FUNCTION_BLOCK GiveWorkpiece (* Composite Function Block Type *)
  (* Standard: 61499-2 *)
  (* Version 0.0, 7/2/2026, template *)
  PACKAGE Main;
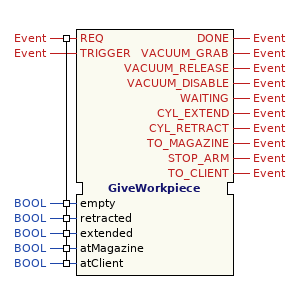
  EVENT_INPUT
    REQ WITH empty, retracted, extended, atMagazine, atClient; (* Normal Execution Request *)
    TRIGGER;
  END_EVENT
  EVENT_OUTPUT
    DONE;
    VACUUM_GRAB;
    VACUUM_RELEASE;
    VACUUM_DISABLE;
    WAITING;
    CYL_EXTEND;
    CYL_RETRACT;
    TO_MAGAZINE;
    STOP_ARM;
    TO_CLIENT;
  END_EVENT
  VAR_INPUT
    empty : BOOL; (* Input event qualifier *)
    retracted : BOOL;
    extended : BOOL;
    atMagazine : BOOL;
    atClient : BOOL;
  END_VAR
  FBS
    FB1 : MagazineSupplyWp;
    ToMagazine : SimpleMove;
    Grab : VacuumSequence;
    ToClient : SimpleMove;
    Release : VacuumSequence;
    FB6 : ArmReset;
    FB7 : E_MERGE;
    FB8 : E_MERGE;
    FB9 : E_MERGE;
    FB10 : E_MERGE;
    FB11 : E_MERGE;
    FB12 : E_MERGE;
  END_FBS
  EVENT_CONNECTIONS
    REQ TO FB1.E7ACA3FA6937DBD5;
    REQ TO ToMagazine.08A6921781769002;
    REQ TO ToClient.08A6921781769002;
    REQ TO FB6.78E8E2AA9DAF29A8;
    TRIGGER TO FB1.CCDC0F1EC03E3A5A;
    FB1.FFF627DF72AA63EC TO CYL_EXTEND;
    FB1.CD1413F90346ACAE TO CYL_RETRACT;
    FB1.F53F7251A3029812 TO ToMagazine.BEEA5224F96B4EAA;
    FB1.C1D84DB1B6EB4247 TO WAITING;
    ToMagazine.19B414802953B8F9 TO Grab.E95F52AEE292CFEA;
    ToMagazine.4A40729E5CEB7782 TO FB11.EI1;
    ToMagazine.FCE01ED48ED44FD9 TO FB12.EI1;
    Grab.8B550AE5A1007C15 TO ToClient.BEEA5224F96B4EAA;
    Grab.5305E856C95E0A15 TO FB7.EI1;
    Grab.2E956B9A6CBDEE5C TO FB8.EI1;
    Grab.993B0E497578A534 TO FB9.EI1;
    ToClient.19B414802953B8F9 TO Release.98EBB230BBACE9D4;
    ToClient.4A40729E5CEB7782 TO FB10.EI1;
    ToClient.FCE01ED48ED44FD9 TO FB12.EI2;
    Release.993B0E497578A534 TO FB9.EI2;
    Release.2E956B9A6CBDEE5C TO FB8.EI2;
    Release.5305E856C95E0A15 TO FB7.EI2;
    Release.8B550AE5A1007C15 TO FB6.44541FA90B36D44F;
    FB6.6B9B16A5CCCF0A5F TO DONE;
    FB6.AF051DE6AC146B46 TO FB10.EI2;
    FB6.88EB222F28F57D09 TO FB11.EI2;
    FB6.4279AF5F2D571F35 TO FB12.EI1;
    FB12.EO TO STOP_ARM;
    FB11.EO TO TO_MAGAZINE;
    FB10.EO TO TO_CLIENT;
    FB9.EO TO VACUUM_DISABLE;
    FB8.EO TO VACUUM_RELEASE;
    FB7.EO TO VACUUM_GRAB;
  END_CONNECTIONS
  DATA_CONNECTIONS
    empty TO FB1.65B96A6108347471;
    retracted TO FB1.F3A16FF43FB1E09C;
    extended TO FB1.F24DAEB350B1D1C4;
    atMagazine TO ToMagazine.D7113296D1A5E867;
    atMagazine TO FB6.4929591747EB6C68;
    atClient TO ToClient.D7113296D1A5E867;
    atClient TO FB6.C845A2BE94918BBD;
  END_CONNECTIONS
END_FUNCTION_BLOCK
